ADAPTER WagoRegCom (* Register communication for Wago modules *)
  (* Standard: 61499-2; Description: Copyright (c) 2026 Monika Wenger This program and the accompanying materials are made available under the terms of the Eclipse Public License 2.0 which is available at https://www.eclipse.org/legal/epl-2.0/ SPDX-License-Identifier: EPL-2.0 *)
  (* Version 3.0, 2026-07-21, Monika Wenger *)
  PACKAGE eclipse4diac::io::wago;
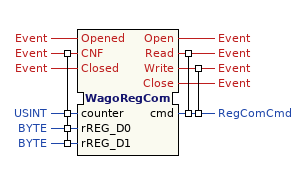
  EVENT_INPUT
    Opened; (* Confirms opening of register communication *)
    CNF WITH counter, rREG_D0, rREG_D1; (* Confirms that the R/W command has been processed *)
    Closed; (* Confirms closing of register communication *)
  END_EVENT
  EVENT_OUTPUT
    Open; (* Open register communication *)
    Read WITH cmd; (* Read register with RegNr *)
    Write WITH cmd; (* Write register with RegNr *)
    Close; (* Close register communication *)
  END_EVENT
  VAR_INPUT
    counter : USINT; (* Counts the commands processed *)
    rREG_D0 : BYTE; (* LSB data read from the register RegNr *)
    rREG_D1 : BYTE; (* MSB data read from the register RegNr *)
  END_VAR
  VAR_OUTPUT
    cmd : eclipse4diac::io::wago::RegComCmd; (* Command for register communication *)
  END_VAR
END_ADAPTER
